(* IEC 61131-3 sources: plc-iiot-stack/tools/tests/fixtures/lowering/src/POUs/FB_Alarm, 2 files *)

(* ---- FB_Alarm.decl.st ---- *)
// Назначение: пример для понижения iec-checker (tools/tests/test_assemble.py)
// Автор:      kr0nsch
// Версия:     0.1.0
// Документ:   docs/LAYOUT.md, раздел «Собранный текст build/assembled»; tools/README.md
FUNCTION_BLOCK FB_Alarm IMPLEMENTS I_Alarm
VAR_INPUT
    xOn : BOOL;
END_VAR
VAR
    iPriority : INT := 1;
    tStamp : TIME;
    ltStamp : LTIME;
    tLimit : TIME := T#1h500ms;
    ltLimit : LTIME := LTIME#1H500MS;
END_VAR

(* ---- FB_Alarm.impl.st ---- *)
// Системное время, длительности с пропуском единиц, пустые операторы и ветви
IF xOn THEN
    tStamp := TIME();
    ltStamp := LTIME();
ELSIF tStamp > t#5s THEN
    ;
ELSE
    // состояние не меняется
END_IF
if tStamp >= T#1h_30m then
    tStamp := tLimit;
end_if;;
